MOVC C01856 V=12.0 ACC=20 DEC=20
MOVC C01857 V=12.0 ACC=20 DEC=20
MOVC C01858 V=12.0 ACC=20 DEC=20
MOVL C01859 V=7.0 ACC=20 DEC=20
MOVL C01860 V=7.0 ACC=20 DEC=20
MOVL C01861 V=7.0 ACC=20 DEC=20
MOVL C01862 V=7.0 ACC=20 DEC=20
MOVL C01863 V=7.0 ACC=20 DEC=20
MOVL C01864 V=7.0 ACC=20 DEC=20
MOVL C01865 V=7.0 ACC=20 DEC=20
MOVL C01866 V=7.0 ACC=20 DEC=20
MOVL C01867 V=7.0 ACC=20 DEC=20
MOVL C01868 V=7.0 PL=1
MOVL C01869 V=7.0 ACC=20 DEC=20
MOVL C01870 V=7.0 ACC=20 DEC=20
MOVL C01871 V=7.0 ACC=20 DEC=20
MOVL C01872 V=7.0 ACC=20 DEC=20
MOVL C01873 V=7.0 ACC=20 DEC=20
MOVL C01874 V=7.0 ACC=20 DEC=20
MOVL C01875 V=7.0 ACC=20 DEC=20
MOVL C01876 V=7.0 ACC=20 DEC=20
MOVL C01877 V=7.0 ACC=20 DEC=20
MOVL C01878 V=7.0 ACC=20 DEC=20
MOVL C01879 V=7.0 ACC=20 DEC=20
MOVL C01880 V=7.0 ACC=20 DEC=20
MOVL C01881 V=7.0 ACC=20 DEC=20
MOVL C01882 V=7.0 ACC=20 DEC=20
MOVL C01883 V=7.0 ACC=20 DEC=20
MOVL C01884 V=7.0 ACC=20 DEC=20
MOVL C01885 V=7.0 ACC=20 DEC=20
MOVL C01886 V=7.0 ACC=20 DEC=20
MOVL C01887 V=7.0 ACC=20 DEC=20
MOVL C01888 V=7.0 ACC=20 DEC=20
MOVL C01889 V=7.0 ACC=20 DEC=20
MOVL C01890 V=7.0 PL=1
MOVL C01891 V=7.0 ACC=20 DEC=20
MOVL C01892 V=7.0 ACC=20 DEC=20
MOVL C01893 V=7.0 ACC=20 DEC=20
MOVL C01894 V=7.0 ACC=20 DEC=20
MOVL C01895 V=7.0 ACC=20 DEC=20
MOVL C01896 V=7.0 ACC=20 DEC=20
MOVL C01897 V=7.0 ACC=20 DEC=20
MOVL C01898 V=7.0 ACC=20 DEC=20
MOVL C01899 V=7.0 ACC=20 DEC=20
MOVC C01900 V=12.0 ACC=20 DEC=20
MOVC C01901 V=12.0 ACC=20 DEC=20
MOVC C01902 V=12.0 ACC=20 DEC=20
MOVL C01903 V=7.0 ACC=20 DEC=20
MOVL C01904 V=7.0 ACC=20 DEC=20
MOVL C01905 V=7.0 ACC=20 DEC=20
MOVL C01906 V=7.0 ACC=20 DEC=20
MOVL C01907 V=7.0 ACC=20 DEC=20
MOVL C01908 V=7.0 ACC=20 DEC=20
MOVL C01909 V=7.0 ACC=20 DEC=20
MOVL C01910 V=7.0 ACC=20 DEC=20
MOVL C01911 V=7.0 ACC=20 DEC=20
MOVL C01912 V=7.0 ACC=20 DEC=20
MOVL C01913 V=7.0 ACC=20 DEC=20
MOVL C01914 V=7.0 ACC=20 DEC=20
MOVL C01915 V=7.0 ACC=20 DEC=20
MOVL C01916 V=7.0 ACC=20 DEC=20
MOVL C01917 V=7.0 ACC=20 DEC=20
MOVL C01918 V=7.0 ACC=20 DEC=20
MOVL C01919 V=7.0 ACC=20 DEC=20
MOVL C01920 V=7.0 ACC=20 DEC=20
MOVL C01921 V=7.0 ACC=20 DEC=20
MOVC C01922 V=12.0 ACC=20 DEC=20
MOVC C01923 V=12.0 ACC=20 DEC=20
MOVC C01924 V=12.0 ACC=20 DEC=20
MOVL C01925 V=7.0 ACC=20 DEC=20
MOVL C01926 V=7.0 ACC=20 DEC=20
MOVL C01927 V=7.0 ACC=20 DEC=20
MOVL C01928 V=7.0 ACC=20 DEC=20
MOVL C01929 V=7.0 ACC=20 DEC=20
MOVL C01930 V=7.0 ACC=20 DEC=20
MOVL C01931 V=7.0 ACC=20 DEC=20
MOVL C01932 V=7.0 ACC=20 DEC=20
MOVL C01933 V=7.0 ACC=20 DEC=20
MOVL C01934 V=7.0 PL=1
MOVL C01935 V=7.0 ACC=20 DEC=20
MOVL C01936 V=7.0 ACC=20 DEC=20
MOVL C01937 V=7.0 ACC=20 DEC=20
MOVL C01938 V=7.0 ACC=20 DEC=20
MOVL C01939 V=7.0 ACC=20 DEC=20
MOVL C01940 V=7.0 ACC=20 DEC=20
MOVL C01941 V=7.0 ACC=20 DEC=20
MOVL C01942 V=7.0 ACC=20 DEC=20
MOVL C01943 V=7.0 ACC=20 DEC=20
MOVL C01944 V=7.0 ACC=20 DEC=20
MOVL C01945 V=7.0 ACC=20 DEC=20
MOVL C01946 V=7.0 ACC=20 DEC=20
MOVL C01947 V=7.0 ACC=20 DEC=20
MOVL C01948 V=7.0 ACC=20 DEC=20
MOVL C01949 V=7.0 ACC=20 DEC=20
MOVL C01950 V=7.0 ACC=20 DEC=20
MOVL C01951 V=7.0 ACC=20 DEC=20
MOVL C01952 V=7.0 ACC=20 DEC=20
MOVL C01953 V=7.0 ACC=20 DEC=20
MOVL C01954 V=7.0 ACC=20 DEC=20
MOVL C01955 V=7.0 ACC=20 DEC=20
MOVL C01956 V=7.0 PL=1
MOVL C01957 V=7.0 ACC=20 DEC=20
MOVL C01958 V=7.0 ACC=20 DEC=20
MOVL C01959 V=7.0 ACC=20 DEC=20
MOVL C01960 V=7.0 ACC=20 DEC=20
MOVL C01961 V=7.0 ACC=20 DEC=20
MOVL C01962 V=7.0 ACC=20 DEC=20
MOVL C01963 V=7.0 ACC=20 DEC=20
MOVL C01964 V=7.0 ACC=20 DEC=20
MOVL C01965 V=7.0 ACC=20 DEC=20
MOVL C01966 V=7.0 ACC=20 DEC=20
ARCOF
TIMER T=30
MOVL C01967 V=11.0 ACC=20 DEC=20
*LAG16
MACRO1 MJ#(0) ARGF2
ARCON
MOVL C01968 V=7.0 ACC=20 DEC=20
MOVL C01969 V=7.0 ACC=20 DEC=20
MOVL C01970 V=7.0 ACC=20 DEC=20
MOVL C01971 V=7.0 ACC=20 DEC=20
MOVL C01972 V=7.0 ACC=20 DEC=20
MOVL C01973 V=7.0 ACC=20 DEC=20
MOVL C01974 V=7.0 ACC=20 DEC=20
MOVL C01975 V=7.0 ACC=20 DEC=20
MOVL C01976 V=7.0 ACC=20 DEC=20
MOVL C01977 V=7.0 PL=1
MOVL C01978 V=7.0 ACC=20 DEC=20
MOVL C01979 V=7.0 ACC=20 DEC=20
MOVL C01980 V=7.0 ACC=20 DEC=20
MOVL C01981 V=7.0 ACC=20 DEC=20
MOVL C01982 V=7.0 ACC=20 DEC=20
MOVL C01983 V=7.0 ACC=20 DEC=20
MOVL C01984 V=7.0 ACC=20 DEC=20
MOVL C01985 V=7.0 ACC=20 DEC=20
MOVL C01986 V=7.0 ACC=20 DEC=20
MOVL C01987 V=7.0 ACC=20 DEC=20
MOVL C01988 V=7.0 ACC=20 DEC=20
MOVL C01989 V=7.0 ACC=20 DEC=20
MOVL C01990 V=7.0 ACC=20 DEC=20
MOVL C01991 V=7.0 ACC=20 DEC=20
MOVL C01992 V=7.0 ACC=20 DEC=20
MOVL C01993 V=7.0 ACC=20 DEC=20
MOVL C01994 V=7.0 ACC=20 DEC=20
MOVL C01995 V=7.0 ACC=20 DEC=20
MOVL C01996 V=7.0 ACC=20 DEC=20
MOVL C01997 V=7.0 ACC=20 DEC=20
MOVL C01998 V=7.0 ACC=20 DEC=20
MOVL C01999 V=7.0 PL=1
MOVL C02000 V=7.0 ACC=20 DEC=20
MOVL C02001 V=7.0 ACC=20 DEC=20
MOVL C02002 V=7.0 ACC=20 DEC=20
MOVL C02003 V=7.0 ACC=20 DEC=20
MOVL C02004 V=7.0 ACC=20 DEC=20
MOVL C02005 V=7.0 ACC=20 DEC=20
MOVL C02006 V=7.0 ACC=20 DEC=20
MOVL C02007 V=7.0 ACC=20 DEC=20
MOVL C02008 V=7.0 ACC=20 DEC=20
MOVC C02009 V=12.0 ACC=20 DEC=20
MOVC C02010 V=12.0 ACC=20 DEC=20
MOVC C02011 V=12.0 ACC=20 DEC=20
MOVL C02012 V=7.0 ACC=20 DEC=20
MOVL C02013 V=7.0 ACC=20 DEC=20
MOVL C02014 V=7.0 ACC=20 DEC=20
MOVL C02015 V=7.0 ACC=20 DEC=20
MOVL C02016 V=7.0 ACC=20 DEC=20
MOVL C02017 V=7.0 ACC=20 DEC=20
MOVL C02018 V=7.0 ACC=20 DEC=20
MOVL C02019 V=7.0 ACC=20 DEC=20
MOVL C02020 V=7.0 ACC=20 DEC=20
MOVL C02021 V=7.0 ACC=20 DEC=20
MOVL C02022 V=7.0 ACC=20 DEC=20
MOVL C02023 V=7.0 ACC=20 DEC=20
MOVL C02024 V=7.0 ACC=20 DEC=20
MOVL C02025 V=7.0 ACC=20 DEC=20
MOVL C02026 V=7.0 ACC=20 DEC=20
MOVL C02027 V=7.0 ACC=20 DEC=20
MOVL C02028 V=7.0 ACC=20 DEC=20
MOVL C02029 V=7.0 ACC=20 DEC=20
MOVL C02030 V=7.0 ACC=20 DEC=20
MOVC C02031 V=12.0 ACC=20 DEC=20
MOVC C02032 V=12.0 ACC=20 DEC=20
MOVC C02033 V=12.0 ACC=20 DEC=20
MOVL C02034 V=7.0 ACC=20 DEC=20
MOVL C02035 V=7.0 ACC=20 DEC=20
MOVL C02036 V=7.0 ACC=20 DEC=20
MOVL C02037 V=7.0 ACC=20 DEC=20
MOVL C02038 V=7.0 ACC=20 DEC=20
MOVL C02039 V=7.0 ACC=20 DEC=20
MOVL C02040 V=7.0 ACC=20 DEC=20
MOVL C02041 V=7.0 ACC=20 DEC=20
MOVL C02042 V=7.0 ACC=20 DEC=20
MOVL C02043 V=7.0 PL=1
MOVL C02044 V=7.0 ACC=20 DEC=20
MOVL C02045 V=7.0 ACC=20 DEC=20
MOVL C02046 V=7.0 ACC=20 DEC=20
MOVL C02047 V=7.0 ACC=20 DEC=20
MOVL C02048 V=7.0 ACC=20 DEC=20
MOVL C02049 V=7.0 ACC=20 DEC=20
MOVL C02050 V=7.0 ACC=20 DEC=20
MOVL C02051 V=7.0 ACC=20 DEC=20
MOVL C02052 V=7.0 ACC=20 DEC=20
MOVL C02053 V=7.0 ACC=20 DEC=20
MOVL C02054 V=7.0 ACC=20 DEC=20
MOVL C02055 V=7.0 ACC=20 DEC=20
MOVL C02056 V=7.0 ACC=20 DEC=20
MOVL C02057 V=7.0 ACC=20 DEC=20
MOVL C02058 V=7.0 ACC=20 DEC=20
MOVL C02059 V=7.0 ACC=20 DEC=20
MOVL C02060 V=7.0 ACC=20 DEC=20
MOVL C02061 V=7.0 ACC=20 DEC=20
MOVL C02062 V=7.0 ACC=20 DEC=20
MOVL C02063 V=7.0 ACC=20 DEC=20
MOVL C02064 V=7.0 ACC=20 DEC=20
MOVL C02065 V=7.0 PL=1
MOVL C02066 V=7.0 ACC=20 DEC=20
MOVL C02067 V=7.0 ACC=20 DEC=20
MOVL C02068 V=7.0 ACC=20 DEC=20
MOVL C02069 V=7.0 ACC=20 DEC=20
MOVL C02070 V=7.0 ACC=20 DEC=20
MOVL C02071 V=7.0 ACC=20 DEC=20
MOVL C02072 V=7.0 ACC=20 DEC=20
MOVL C02073 V=7.0 ACC=20 DEC=20
MOVL C02074 V=7.0 ACC=20 DEC=20
MOVC C02075 V=12.0 ACC=20 DEC=20
MOVC C02076 V=12.0 ACC=20 DEC=20
MOVC C02077 V=12.0 ACC=20 DEC=20
MOVL C02078 V=7.0 ACC=20 DEC=20
MOVL C02079 V=7.0 ACC=20 DEC=20
MOVL C02080 V=7.0 ACC=20 DEC=20
MOVL C02081 V=7.0 ACC=20 DEC=20
MOVL C02082 V=7.0 ACC=20 DEC=20
MOVL C02083 V=7.0 ACC=20 DEC=20
MOVL C02084 V=7.0 ACC=20 DEC=20
MOVL C02085 V=7.0 ACC=20 DEC=20
MOVL C02086 V=7.0 ACC=20 DEC=20
MOVL C02087 V=7.0 ACC=20 DEC=20
MOVL C02088 V=7.0 ACC=20 DEC=20
MOVL C02089 V=7.0 ACC=20 DEC=20
MOVL C02090 V=7.0 ACC=20 DEC=20
MOVL C02091 V=7.0 ACC=20 DEC=20
MOVL C02092 V=7.0 ACC=20 DEC=20
MOVL C02093 V=7.0 ACC=20 DEC=20
MOVL C02094 V=7.0 ACC=20 DEC=20
MOVL C02095 V=7.0 ACC=20 DEC=20
MOVL C02096 V=7.0 ACC=20 DEC=20
MOVL C02097 V=7.0 ACC=20 DEC=20
ARCOF
TIMER T=30
MOVL C02098 V=11.0 ACC=20 DEC=20
*LAG17
MACRO1 MJ#(0) ARGF2
ARCON
MOVL C02099 V=7.0 ACC=20 DEC=20
MOVL C02100 V=7.0 ACC=20 DEC=20
MOVL C02101 V=7.0 ACC=20 DEC=20
MOVL C02102 V=7.0 ACC=20 DEC=20
MOVL C02103 V=7.0 ACC=20 DEC=20
MOVL C02104 V=7.0 ACC=20 DEC=20
MOVL C02105 V=7.0 ACC=20 DEC=20
MOVL C02106 V=7.0 ACC=20 DEC=20
MOVL C02107 V=7.0 ACC=20 DEC=20
MOVL C02108 V=7.0 ACC=20 DEC=20
MOVL C02109 V=7.0 ACC=20 DEC=20
MOVL C02110 V=7.0 ACC=20 DEC=20
MOVL C02111 V=7.0 ACC=20 DEC=20
MOVL C02112 V=7.0 ACC=20 DEC=20
MOVL C02113 V=7.0 ACC=20 DEC=20
MOVL C02114 V=7.0 ACC=20 DEC=20
MOVL C02115 V=7.0 ACC=20 DEC=20
MOVL C02116 V=7.0 ACC=20 DEC=20
MOVL C02117 V=7.0 ACC=20 DEC=20
MOVC C02118 V=12.0 ACC=20 DEC=20
MOVC C02119 V=12.0 ACC=20 DEC=20
MOVC C02120 V=12.0 ACC=20 DEC=20
MOVL C02121 V=7.0 ACC=20 DEC=20
MOVL C02122 V=7.0 ACC=20 DEC=20
MOVL C02123 V=7.0 ACC=20 DEC=20
MOVL C02124 V=7.0 ACC=20 DEC=20
MOVL C02125 V=7.0 ACC=20 DEC=20
MOVL C02126 V=7.0 ACC=20 DEC=20
MOVL C02127 V=7.0 ACC=20 DEC=20
MOVL C02128 V=7.0 ACC=20 DEC=20
MOVL C02129 V=7.0 ACC=20 DEC=20
MOVL C02130 V=7.0 PL=1
MOVL C02131 V=7.0 ACC=20 DEC=20
MOVL C02132 V=7.0 ACC=20 DEC=20
MOVL C02133 V=7.0 ACC=20 DEC=20
MOVL C02134 V=7.0 ACC=20 DEC=20
MOVL C02135 V=7.0 ACC=20 DEC=20
MOVL C02136 V=7.0 ACC=20 DEC=20
MOVL C02137 V=7.0 ACC=20 DEC=20
MOVL C02138 V=7.0 ACC=20 DEC=20
MOVL C02139 V=7.0 ACC=20 DEC=20
MOVL C02140 V=7.0 ACC=20 DEC=20
MOVL C02141 V=7.0 ACC=20 DEC=20
MOVL C02142 V=7.0 ACC=20 DEC=20
MOVL C02143 V=7.0 ACC=20 DEC=20
MOVL C02144 V=7.0 ACC=20 DEC=20
MOVL C02145 V=7.0 ACC=20 DEC=20
MOVL C02146 V=7.0 ACC=20 DEC=20
MOVL C02147 V=7.0 ACC=20 DEC=20
MOVL C02148 V=7.0 ACC=20 DEC=20
MOVL C02149 V=7.0 ACC=20 DEC=20
MOVL C02150 V=7.0 ACC=20 DEC=20
MOVL C02151 V=7.0 ACC=20 DEC=20
MOVL C02152 V=7.0 PL=1
MOVL C02153 V=7.0 ACC=20 DEC=20
MOVL C02154 V=7.0 ACC=20 DEC=20
MOVL C02155 V=7.0 ACC=20 DEC=20
MOVL C02156 V=7.0 ACC=20 DEC=20
MOVL C02157 V=7.0 ACC=20 DEC=20
MOVL C02158 V=7.0 ACC=20 DEC=20
MOVL C02159 V=7.0 ACC=20 DEC=20
MOVL C02160 V=7.0 ACC=20 DEC=20
MOVL C02161 V=7.0 ACC=20 DEC=20
MOVC C02162 V=12.0 ACC=20 DEC=20
MOVC C02163 V=12.0 ACC=20 DEC=20
MOVC C02164 V=12.0 ACC=20 DEC=20
MOVL C02165 V=7.0 ACC=20 DEC=20
MOVL C02166 V=7.0 ACC=20 DEC=20
MOVL C02167 V=7.0 ACC=20 DEC=20
MOVL C02168 V=7.0 ACC=20 DEC=20
MOVL C02169 V=7.0 ACC=20 DEC=20
MOVL C02170 V=7.0 ACC=20 DEC=20
MOVL C02171 V=7.0 ACC=20 DEC=20
MOVL C02172 V=7.0 ACC=20 DEC=20
MOVL C02173 V=7.0 ACC=20 DEC=20
MOVL C02174 V=7.0 ACC=20 DEC=20
MOVL C02175 V=7.0 ACC=20 DEC=20
MOVL C02176 V=7.0 ACC=20 DEC=20
MOVL C02177 V=7.0 ACC=20 DEC=20
MOVL C02178 V=7.0 ACC=20 DEC=20
MOVL C02179 V=7.0 ACC=20 DEC=20
MOVL C02180 V=7.0 ACC=20 DEC=20
MOVL C02181 V=7.0 ACC=20 DEC=20
MOVL C02182 V=7.0 ACC=20 DEC=20
MOVL C02183 V=7.0 ACC=20 DEC=20
MOVC C02184 V=12.0 ACC=20 DEC=20
MOVC C02185 V=12.0 ACC=20 DEC=20
MOVC C02186 V=12.0 ACC=20 DEC=20
MOVL C02187 V=7.0 ACC=20 DEC=20
MOVL C02188 V=7.0 ACC=20 DEC=20
MOVL C02189 V=7.0 ACC=20 DEC=20
MOVL C02190 V=7.0 ACC=20 DEC=20
MOVL C02191 V=7.0 ACC=20 DEC=20
MOVL C02192 V=7.0 ACC=20 DEC=20
MOVL C02193 V=7.0 ACC=20 DEC=20
MOVL C02194 V=7.0 ACC=20 DEC=20
MOVL C02195 V=7.0 ACC=20 DEC=20
MOVL C02196 V=7.0 PL=1
MOVL C02197 V=7.0 ACC=20 DEC=20
MOVL C02198 V=7.0 ACC=20 DEC=20
MOVL C02199 V=7.0 ACC=20 DEC=20
MOVL C02200 V=7.0 ACC=20 DEC=20
MOVL C02201 V=7.0 ACC=20 DEC=20
MOVL C02202 V=7.0 ACC=20 DEC=20
MOVL C02203 V=7.0 ACC=20 DEC=20
MOVL C02204 V=7.0 ACC=20 DEC=20
MOVL C02205 V=7.0 ACC=20 DEC=20
MOVL C02206 V=7.0 ACC=20 DEC=20
MOVL C02207 V=7.0 ACC=20 DEC=20
MOVL C02208 V=7.0 ACC=20 DEC=20
MOVL C02209 V=7.0 ACC=20 DEC=20
MOVL C02210 V=7.0 ACC=20 DEC=20
MOVL C02211 V=7.0 ACC=20 DEC=20
MOVL C02212 V=7.0 ACC=20 DEC=20
MOVL C02213 V=7.0 ACC=20 DEC=20
MOVL C02214 V=7.0 ACC=20 DEC=20
MOVL C02215 V=7.0 ACC=20 DEC=20
MOVL C02216 V=7.0 ACC=20 DEC=20
MOVL C02217 V=7.0 ACC=20 DEC=20
MOVL C02218 V=7.0 PL=1
MOVL C02219 V=7.0 ACC=20 DEC=20
MOVL C02220 V=7.0 ACC=20 DEC=20
MOVL C02221 V=7.0 ACC=20 DEC=20
MOVL C02222 V=7.0 ACC=20 DEC=20
MOVL C02223 V=7.0 ACC=20 DEC=20
MOVL C02224 V=7.0 ACC=20 DEC=20
MOVL C02225 V=7.0 ACC=20 DEC=20
MOVL C02226 V=7.0 ACC=20 DEC=20
MOVL C02227 V=7.0 ACC=20 DEC=20
MOVL C02228 V=7.0 ACC=20 DEC=20
ARCOF
TIMER T=30
MOVL C02229 V=11.0 ACC=20 DEC=20
*LAG18
MACRO1 MJ#(0) ARGF2
ARCON
MOVL C02230 V=7.0 ACC=20 DEC=20
MOVL C02231 V=7.0 ACC=20 DEC=20
MOVL C02232 V=7.0 ACC=20 DEC=20
MOVL C02233 V=7.0 ACC=20 DEC=20
MOVL C02234 V=7.0 ACC=20 DEC=20
MOVL C02235 V=7.0 ACC=20 DEC=20
MOVL C02236 V=7.0 ACC=20 DEC=20
MOVL C02237 V=7.0 ACC=20 DEC=20
MOVL C02238 V=7.0 ACC=20 DEC=20
MOVL C02239 V=7.0 PL=1
MOVL C02240 V=7.0 ACC=20 DEC=20
MOVL C02241 V=7.0 ACC=20 DEC=20
MOVL C02242 V=7.0 ACC=20 DEC=20
MOVL C02243 V=7.0 ACC=20 DEC=20
MOVL C02244 V=7.0 ACC=20 DEC=20
MOVL C02245 V=7.0 ACC=20 DEC=20
MOVL C02246 V=7.0 ACC=20 DEC=20
MOVL C02247 V=7.0 ACC=20 DEC=20
MOVL C02248 V=7.0 ACC=20 DEC=20
MOVL C02249 V=7.0 ACC=20 DEC=20
MOVL C02250 V=7.0 ACC=20 DEC=20
MOVL C02251 V=7.0 ACC=20 DEC=20
MOVL C02252 V=7.0 ACC=20 DEC=20
MOVL C02253 V=7.0 ACC=20 DEC=20
MOVL C02254 V=7.0 ACC=20 DEC=20
MOVL C02255 V=7.0 ACC=20 DEC=20
MOVL C02256 V=7.0 ACC=20 DEC=20
MOVL C02257 V=7.0 ACC=20 DEC=20
MOVL C02258 V=7.0 ACC=20 DEC=20
MOVL C02259 V=7.0 ACC=20 DEC=20
MOVL C02260 V=7.0 ACC=20 DEC=20
MOVL C02261 V=7.0 PL=1
MOVL C02262 V=7.0 ACC=20 DEC=20
MOVL C02263 V=7.0 ACC=20 DEC=20
MOVL C02264 V=7.0 ACC=20 DEC=20
MOVL C02265 V=7.0 ACC=20 DEC=20
MOVL C02266 V=7.0 ACC=20 DEC=20
MOVL C02267 V=7.0 ACC=20 DEC=20
MOVL C02268 V=7.0 ACC=20 DEC=20
MOVL C02269 V=7.0 ACC=20 DEC=20
MOVL C02270 V=7.0 ACC=20 DEC=20
MOVC C02271 V=12.0 ACC=20 DEC=20
MOVC C02272 V=12.0 ACC=20 DEC=20
MOVC C02273 V=12.0 ACC=20 DEC=20
MOVL C02274 V=7.0 ACC=20 DEC=20
MOVL C02275 V=7.0 ACC=20 DEC=20
MOVL C02276 V=7.0 ACC=20 DEC=20
MOVL C02277 V=7.0 ACC=20 DEC=20
MOVL C02278 V=7.0 ACC=20 DEC=20
MOVL C02279 V=7.0 ACC=20 DEC=20
MOVL C02280 V=7.0 ACC=20 DEC=20
MOVL C02281 V=7.0 ACC=20 DEC=20
MOVL C02282 V=7.0 ACC=20 DEC=20
MOVL C02283 V=7.0 ACC=20 DEC=20
MOVL C02284 V=7.0 ACC=20 DEC=20
MOVL C02285 V=7.0 ACC=20 DEC=20
MOVL C02286 V=7.0 ACC=20 DEC=20
MOVL C02287 V=7.0 ACC=20 DEC=20
MOVL C02288 V=7.0 ACC=20 DEC=20
MOVL C02289 V=7.0 ACC=20 DEC=20
MOVL C02290 V=7.0 ACC=20 DEC=20
MOVL C02291 V=7.0 ACC=20 DEC=20
MOVL C02292 V=7.0 ACC=20 DEC=20
MOVC C02293 V=12.0 ACC=20 DEC=20
MOVC C02294 V=12.0 ACC=20 DEC=20
MOVC C02295 V=12.0 ACC=20 DEC=20
MOVL C02296 V=7.0 ACC=20 DEC=20
MOVL C02297 V=7.0 ACC=20 DEC=20
MOVL C02298 V=7.0 ACC=20 DEC=20
MOVL C02299 V=7.0 ACC=20 DEC=20
MOVL C02300 V=7.0 ACC=20 DEC=20
MOVL C02301 V=7.0 ACC=20 DEC=20
MOVL C02302 V=7.0 ACC=20 DEC=20
MOVL C02303 V=7.0 ACC=20 DEC=20
MOVL C02304 V=7.0 ACC=20 DEC=20
MOVL C02305 V=7.0 PL=1
MOVL C02306 V=7.0 ACC=20 DEC=20
MOVL C02307 V=7.0 ACC=20 DEC=20
MOVL C02308 V=7.0 ACC=20 DEC=20
MOVL C02309 V=7.0 ACC=20 DEC=20
MOVL C02310 V=7.0 ACC=20 DEC=20
MOVL C02311 V=7.0 ACC=20 DEC=20
MOVL C02312 V=7.0 ACC=20 DEC=20
MOVL C02313 V=7.0 ACC=20 DEC=20
MOVL C02314 V=7.0 ACC=20 DEC=20
MOVL C02315 V=7.0 ACC=20 DEC=20
MOVL C02316 V=7.0 ACC=20 DEC=20
MOVL C02317 V=7.0 ACC=20 DEC=20
MOVL C02318 V=7.0 ACC=20 DEC=20
MOVL C02319 V=7.0 ACC=20 DEC=20
MOVL C02320 V=7.0 ACC=20 DEC=20
MOVL C02321 V=7.0 ACC=20 DEC=20
MOVL C02322 V=7.0 ACC=20 DEC=20
MOVL C02323 V=7.0 ACC=20 DEC=20
MOVL C02324 V=7.0 ACC=20 DEC=20
MOVL C02325 V=7.0 ACC=20 DEC=20
MOVL C02326 V=7.0 ACC=20 DEC=20
MOVL C02327 V=7.0 PL=1
MOVL C02328 V=7.0 ACC=20 DEC=20
MOVL C02329 V=7.0 ACC=20 DEC=20
MOVL C02330 V=7.0 ACC=20 DEC=20
MOVL C02331 V=7.0 ACC=20 DEC=20
MOVL C02332 V=7.0 ACC=20 DEC=20
MOVL C02333 V=7.0 ACC=20 DEC=20
MOVL C02334 V=7.0 ACC=20 DEC=20
MOVL C02335 V=7.0 ACC=20 DEC=20
MOVL C02336 V=7.0 ACC=20 DEC=20
MOVC C02337 V=12.0 ACC=20 DEC=20
MOVC C02338 V=12.0 ACC=20 DEC=20
MOVC C02339 V=12.0 ACC=20 DEC=20
MOVL C02340 V=7.0 ACC=20 DEC=20
MOVL C02341 V=7.0 ACC=20 DEC=20
MOVL C02342 V=7.0 ACC=20 DEC=20
MOVL C02343 V=7.0 ACC=20 DEC=20
MOVL C02344 V=7.0 ACC=20 DEC=20
MOVL C02345 V=7.0 ACC=20 DEC=20
MOVL C02346 V=7.0 ACC=20 DEC=20
MOVL C02347 V=7.0 ACC=20 DEC=20
MOVL C02348 V=7.0 ACC=20 DEC=20
MOVL C02349 V=7.0 ACC=20 DEC=20
MOVL C02350 V=7.0 ACC=20 DEC=20
MOVL C02351 V=7.0 ACC=20 DEC=20
MOVL C02352 V=7.0 ACC=20 DEC=20
MOVL C02353 V=7.0 ACC=20 DEC=20
MOVL C02354 V=7.0 ACC=20 DEC=20
MOVL C02355 V=7.0 ACC=20 DEC=20
MOVL C02356 V=7.0 ACC=20 DEC=20
MOVL C02357 V=7.0 ACC=20 DEC=20
MOVL C02358 V=7.0 ACC=20 DEC=20
MOVL C02359 V=7.0 ACC=20 DEC=20
ARCOF
TIMER T=30
MOVL C02360 V=11.0 ACC=20 DEC=20
*LAG19
MACRO1 MJ#(0) ARGF2
ARCON
MOVL C02361 V=7.0 ACC=20 DEC=20
MOVL C02362 V=7.0 ACC=20 DEC=20
MOVL C02363 V=7.0 ACC=20 DEC=20
MOVL C02364 V=7.0 ACC=20 DEC=20
MOVL C02365 V=7.0 ACC=20 DEC=20
MOVL C02366 V=7.0 ACC=20 DEC=20
MOVL C02367 V=7.0 ACC=20 DEC=20
MOVL C02368 V=7.0 ACC=20 DEC=20
MOVL C02369 V=7.0 ACC=20 DEC=20
MOVL C02370 V=7.0 ACC=20 DEC=20
MOVL C02371 V=7.0 ACC=20 DEC=20
MOVL C02372 V=7.0 ACC=20 DEC=20
MOVL C02373 V=7.0 ACC=20 DEC=20
MOVL C02374 V=7.0 ACC=20 DEC=20
MOVL C02375 V=7.0 ACC=20 DEC=20
MOVL C02376 V=7.0 ACC=20 DEC=20
MOVL C02377 V=7.0 ACC=20 DEC=20
MOVL C02378 V=7.0 ACC=20 DEC=20
MOVL C02379 V=7.0 ACC=20 DEC=20
MOVC C02380 V=12.0 ACC=20 DEC=20
MOVC C02381 V=12.0 ACC=20 DEC=20
MOVC C02382 V=12.0 ACC=20 DEC=20
MOVL C02383 V=7.0 ACC=20 DEC=20
MOVL C02384 V=7.0 ACC=20 DEC=20
MOVL C02385 V=7.0 ACC=20 DEC=20
MOVL C02386 V=7.0 ACC=20 DEC=20
MOVL C02387 V=7.0 ACC=20 DEC=20
MOVL C02388 V=7.0 ACC=20 DEC=20
MOVL C02389 V=7.0 ACC=20 DEC=20
MOVL C02390 V=7.0 ACC=20 DEC=20
MOVL C02391 V=7.0 ACC=20 DEC=20
MOVL C02392 V=7.0 PL=1
MOVL C02393 V=7.0 ACC=20 DEC=20
MOVL C02394 V=7.0 ACC=20 DEC=20
MOVL C02395 V=7.0 ACC=20 DEC=20
MOVL C02396 V=7.0 ACC=20 DEC=20
MOVL C02397 V=7.0 ACC=20 DEC=20
MOVL C02398 V=7.0 ACC=20 DEC=20
MOVL C02399 V=7.0 ACC=20 DEC=20
MOVL C02400 V=7.0 ACC=20 DEC=20
MOVL C02401 V=7.0 ACC=20 DEC=20
MOVL C02402 V=7.0 ACC=20 DEC=20
MOVL C02403 V=7.0 ACC=20 DEC=20
MOVL C02404 V=7.0 ACC=20 DEC=20
MOVL C02405 V=7.0 ACC=20 DEC=20
MOVL C02406 V=7.0 ACC=20 DEC=20
MOVL C02407 V=7.0 ACC=20 DEC=20
MOVL C02408 V=7.0 ACC=20 DEC=20
MOVL C02409 V=7.0 ACC=20 DEC=20
MOVL C02410 V=7.0 ACC=20 DEC=20
MOVL C02411 V=7.0 ACC=20 DEC=20
MOVL C02412 V=7.0 ACC=20 DEC=20
MOVL C02413 V=7.0 ACC=20 DEC=20
MOVL C02414 V=7.0 PL=1
MOVL C02415 V=7.0 ACC=20 DEC=20
MOVL C02416 V=7.0 ACC=20 DEC=20
MOVL C02417 V=7.0 ACC=20 DEC=20
MOVL C02418 V=7.0 ACC=20 DEC=20
MOVL C02419 V=7.0 ACC=20 DEC=20
MOVL C02420 V=7.0 ACC=20 DEC=20
MOVL C02421 V=7.0 ACC=20 DEC=20
MOVL C02422 V=7.0 ACC=20 DEC=20
MOVL C02423 V=7.0 ACC=20 DEC=20
MOVC C02424 V=12.0 ACC=20 DEC=20
MOVC C02425 V=12.0 ACC=20 DEC=20
MOVC C02426 V=12.0 ACC=20 DEC=20
MOVL C02427 V=7.0 ACC=20 DEC=20
MOVL C02428 V=7.0 ACC=20 DEC=20
MOVL C02429 V=7.0 ACC=20 DEC=20
MOVL C02430 V=7.0 ACC=20 DEC=20
MOVL C02431 V=7.0 ACC=20 DEC=20
MOVL C02432 V=7.0 ACC=20 DEC=20
MOVL C02433 V=7.0 ACC=20 DEC=20
MOVL C02434 V=7.0 ACC=20 DEC=20
MOVL C02435 V=7.0 ACC=20 DEC=20
MOVL C02436 V=7.0 ACC=20 DEC=20
MOVL C02437 V=7.0 ACC=20 DEC=20
MOVL C02438 V=7.0 ACC=20 DEC=20
MOVL C02439 V=7.0 ACC=20 DEC=20
MOVL C02440 V=7.0 ACC=20 DEC=20
MOVL C02441 V=7.0 ACC=20 DEC=20
MOVL C02442 V=7.0 ACC=20 DEC=20
MOVL C02443 V=7.0 ACC=20 DEC=20
MOVL C02444 V=7.0 ACC=20 DEC=20
MOVL C02445 V=7.0 ACC=20 DEC=20
MOVC C02446 V=12.0 ACC=20 DEC=20
MOVC C02447 V=12.0 ACC=20 DEC=20
MOVC C02448 V=12.0 ACC=20 DEC=20
MOVL C02449 V=7.0 ACC=20 DEC=20
MOVL C02450 V=7.0 ACC=20 DEC=20
MOVL C02451 V=7.0 ACC=20 DEC=20
MOVL C02452 V=7.0 ACC=20 DEC=20
MOVL C02453 V=7.0 ACC=20 DEC=20
MOVL C02454 V=7.0 ACC=20 DEC=20
MOVL C02455 V=7.0 ACC=20 DEC=20
MOVL C02456 V=7.0 ACC=20 DEC=20
MOVL C02457 V=7.0 ACC=20 DEC=20
MOVL C02458 V=7.0 PL=1
MOVL C02459 V=7.0 ACC=20 DEC=20
MOVL C02460 V=7.0 ACC=20 DEC=20
MOVL C02461 V=7.0 ACC=20 DEC=20
MOVL C02462 V=7.0 ACC=20 DEC=20
MOVL C02463 V=7.0 ACC=20 DEC=20
MOVL C02464 V=7.0 ACC=20 DEC=20
MOVL C02465 V=7.0 ACC=20 DEC=20
MOVL C02466 V=7.0 ACC=20 DEC=20
MOVL C02467 V=7.0 ACC=20 DEC=20
MOVL C02468 V=7.0 ACC=20 DEC=20
MOVL C02469 V=7.0 ACC=20 DEC=20
MOVL C02470 V=7.0 ACC=20 DEC=20
MOVL C02471 V=7.0 ACC=20 DEC=20
MOVL C02472 V=7.0 ACC=20 DEC=20
MOVL C02473 V=7.0 ACC=20 DEC=20
MOVL C02474 V=7.0 ACC=20 DEC=20
MOVL C02475 V=7.0 ACC=20 DEC=20
MOVL C02476 V=7.0 ACC=20 DEC=20
MOVL C02477 V=7.0 ACC=20 DEC=20
MOVL C02478 V=7.0 ACC=20 DEC=20
MOVL C02479 V=7.0 ACC=20 DEC=20
MOVL C02480 V=7.0 PL=1
MOVL C02481 V=7.0 ACC=20 DEC=20
MOVL C02482 V=7.0 ACC=20 DEC=20
MOVL C02483 V=7.0 ACC=20 DEC=20
MOVL C02484 V=7.0 ACC=20 DEC=20
MOVL C02485 V=7.0 ACC=20 DEC=20
MOVL C02486 V=7.0 ACC=20 DEC=20
MOVL C02487 V=7.0 ACC=20 DEC=20
MOVL C02488 V=7.0 ACC=20 DEC=20
MOVL C02489 V=7.0 ACC=20 DEC=20
MOVL C02490 V=7.0 ACC=20 DEC=20
ARCOF
TIMER T=30
MOVL C02491 V=11.0 ACC=20 DEC=20
*LAG20
MACRO1 MJ#(0) ARGF2
ARCON
MOVL C02492 V=7.0 ACC=20 DEC=20
MOVL C02493 V=7.0 ACC=20 DEC=20
MOVL C02494 V=7.0 ACC=20 DEC=20
MOVL C02495 V=7.0 ACC=20 DEC=20
MOVL C02496 V=7.0 ACC=20 DEC=20
MOVL C02497 V=7.0 ACC=20 DEC=20
MOVL C02498 V=7.0 ACC=20 DEC=20
MOVL C02499 V=7.0 ACC=20 DEC=20
MOVL C02500 V=7.0 ACC=20 DEC=20
MOVL C02501 V=7.0 PL=1
MOVL C02502 V=7.0 ACC=20 DEC=20
MOVL C02503 V=7.0 ACC=20 DEC=20
MOVL C02504 V=7.0 ACC=20 DEC=20
MOVL C02505 V=7.0 ACC=20 DEC=20
MOVL C02506 V=7.0 ACC=20 DEC=20
MOVL C02507 V=7.0 ACC=20 DEC=20
MOVL C02508 V=7.0 ACC=20 DEC=20
MOVL C02509 V=7.0 ACC=20 DEC=20
MOVL C02510 V=7.0 ACC=20 DEC=20
MOVL C02511 V=7.0 ACC=20 DEC=20
MOVL C02512 V=7.0 ACC=20 DEC=20
MOVL C02513 V=7.0 ACC=20 DEC=20
MOVL C02514 V=7.0 ACC=20 DEC=20
MOVL C02515 V=7.0 ACC=20 DEC=20
MOVL C02516 V=7.0 ACC=20 DEC=20
MOVL C02517 V=7.0 ACC=20 DEC=20
MOVL C02518 V=7.0 ACC=20 DEC=20
MOVL C02519 V=7.0 ACC=20 DEC=20
MOVL C02520 V=7.0 ACC=20 DEC=20
MOVL C02521 V=7.0 ACC=20 DEC=20
MOVL C02522 V=7.0 ACC=20 DEC=20
MOVL C02523 V=7.0 PL=1
MOVL C02524 V=7.0 ACC=20 DEC=20
MOVL C02525 V=7.0 ACC=20 DEC=20
MOVL C02526 V=7.0 ACC=20 DEC=20
MOVL C02527 V=7.0 ACC=20 DEC=20
MOVL C02528 V=7.0 ACC=20 DEC=20
MOVL C02529 V=7.0 ACC=20 DEC=20
MOVL C02530 V=7.0 ACC=20 DEC=20
MOVL C02531 V=7.0 ACC=20 DEC=20
MOVL C02532 V=7.0 ACC=20 DEC=20
MOVC C02533 V=12.0 ACC=20 DEC=20
MOVC C02534 V=12.0 ACC=20 DEC=20
MOVC C02535 V=12.0 ACC=20 DEC=20
MOVL C02536 V=7.0 ACC=20 DEC=20
MOVL C02537 V=7.0 ACC=20 DEC=20
MOVL C02538 V=7.0 ACC=20 DEC=20
MOVL C02539 V=7.0 ACC=20 DEC=20
MOVL C02540 V=7.0 ACC=20 DEC=20
MOVL C02541 V=7.0 ACC=20 DEC=20
MOVL C02542 V=7.0 ACC=20 DEC=20
MOVL C02543 V=7.0 ACC=20 DEC=20
MOVL C02544 V=7.0 ACC=20 DEC=20
MOVL C02545 V=7.0 ACC=20 DEC=20
MOVL C02546 V=7.0 ACC=20 DEC=20
MOVL C02547 V=7.0 ACC=20 DEC=20
MOVL C02548 V=7.0 ACC=20 DEC=20
MOVL C02549 V=7.0 ACC=20 DEC=20
MOVL C02550 V=7.0 ACC=20 DEC=20
MOVL C02551 V=7.0 ACC=20 DEC=20
MOVL C02552 V=7.0 ACC=20 DEC=20
MOVL C02553 V=7.0 ACC=20 DEC=20
MOVL C02554 V=7.0 ACC=20 DEC=20
MOVC C02555 V=12.0 ACC=20 DEC=20
MOVC C02556 V=12.0 ACC=20 DEC=20
MOVC C02557 V=12.0 ACC=20 DEC=20
MOVL C02558 V=7.0 ACC=20 DEC=20
MOVL C02559 V=7.0 ACC=20 DEC=20
MOVL C02560 V=7.0 ACC=20 DEC=20
MOVL C02561 V=7.0 ACC=20 DEC=20
MOVL C02562 V=7.0 ACC=20 DEC=20
MOVL C02563 V=7.0 ACC=20 DEC=20
MOVL C02564 V=7.0 ACC=20 DEC=20
MOVL C02565 V=7.0 ACC=20 DEC=20
MOVL C02566 V=7.0 ACC=20 DEC=20
MOVL C02567 V=7.0 PL=1
MOVL C02568 V=7.0 ACC=20 DEC=20
MOVL C02569 V=7.0 ACC=20 DEC=20
MOVL C02570 V=7.0 ACC=20 DEC=20
MOVL C02571 V=7.0 ACC=20 DEC=20
MOVL C02572 V=7.0 ACC=20 DEC=20
MOVL C02573 V=7.0 ACC=20 DEC=20
MOVL C02574 V=7.0 ACC=20 DEC=20
MOVL C02575 V=7.0 ACC=20 DEC=20
MOVL C02576 V=7.0 ACC=20 DEC=20
MOVL C02577 V=7.0 ACC=20 DEC=20
MOVL C02578 V=7.0 ACC=20 DEC=20
MOVL C02579 V=7.0 ACC=20 DEC=20
MOVL C02580 V=7.0 ACC=20 DEC=20
MOVL C02581 V=7.0 ACC=20 DEC=20
MOVL C02582 V=7.0 ACC=20 DEC=20
MOVL C02583 V=7.0 ACC=20 DEC=20
MOVL C02584 V=7.0 ACC=20 DEC=20
MOVL C02585 V=7.0 ACC=20 DEC=20
MOVL C02586 V=7.0 ACC=20 DEC=20
MOVL C02587 V=7.0 ACC=20 DEC=20
MOVL C02588 V=7.0 ACC=20 DEC=20
MOVL C02589 V=7.0 PL=1
MOVL C02590 V=7.0 ACC=20 DEC=20
MOVL C02591 V=7.0 ACC=20 DEC=20
MOVL C02592 V=7.0 ACC=20 DEC=20
MOVL C02593 V=7.0 ACC=20 DEC=20
MOVL C02594 V=7.0 ACC=20 DEC=20
MOVL C02595 V=7.0 ACC=20 DEC=20
MOVL C02596 V=7.0 ACC=20 DEC=20
MOVL C02597 V=7.0 ACC=20 DEC=20
MOVL C02598 V=7.0 ACC=20 DEC=20
MOVC C02599 V=12.0 ACC=20 DEC=20
MOVC C02600 V=12.0 ACC=20 DEC=20
MOVC C02601 V=12.0 ACC=20 DEC=20
MOVL C02602 V=7.0 ACC=20 DEC=20
MOVL C02603 V=7.0 ACC=20 DEC=20
MOVL C02604 V=7.0 ACC=20 DEC=20
MOVL C02605 V=7.0 ACC=20 DEC=20
MOVL C02606 V=7.0 ACC=20 DEC=20
MOVL C02607 V=7.0 ACC=20 DEC=20
MOVL C02608 V=7.0 ACC=20 DEC=20
MOVL C02609 V=7.0 ACC=20 DEC=20
MOVL C02610 V=7.0 ACC=20 DEC=20
MOVL C02611 V=7.0 ACC=20 DEC=20
MOVL C02612 V=7.0 ACC=20 DEC=20
MOVL C02613 V=7.0 ACC=20 DEC=20
MOVL C02614 V=7.0 ACC=20 DEC=20
MOVL C02615 V=7.0 ACC=20 DEC=20
MOVL C02616 V=7.0 ACC=20 DEC=20
MOVL C02617 V=7.0 ACC=20 DEC=20
MOVL C02618 V=7.0 ACC=20 DEC=20
MOVL C02619 V=7.0 ACC=20 DEC=20
MOVL C02620 V=7.0 ACC=20 DEC=20
MOVL C02621 V=7.0 ACC=20 DEC=20
ARCOF
TIMER T=30
MOVL C02622 V=11.0 ACC=20 DEC=20
MOVJ C02623 VJ=0.78
END
